FUNCTION_BLOCK MGZ_IMC (* Extracted Composite Function Block Type *)
  (* Standard: 61499-2 *)
  (* Version 10/20/2026, lizar *)
  PACKAGE Main;
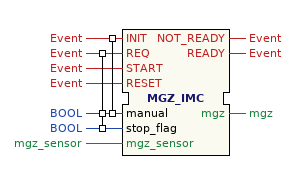
  EVENT_INPUT
    INIT WITH manual; (* Initialization Request *)
    REQ WITH manual, stop_flag; (* Normal Execution Request *)
    START;
    RESET;
  END_EVENT
  EVENT_OUTPUT
    NOT_READY;
    READY;
  END_EVENT
  VAR_INPUT
    manual : BOOL;
    stop_flag : BOOL;
  END_VAR
  SOCKETS
    mgz_sensor : mgz_sensor;
  END_SOCKETS
  PLUGS
    mgz : mgz;
  END_PLUGS
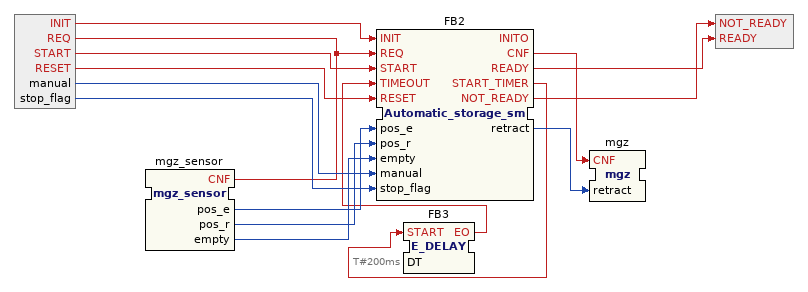
  FBS
    FB2 : Automatic_storage_sm;
    FB3 : E_DELAY(DT := T#200ms);
  END_FBS
  EVENT_CONNECTIONS
    FB2.START_TIMER TO FB3.START;
    FB3.EO TO FB2.TIMEOUT;
    INIT TO FB2.INIT;
    REQ TO FB2.REQ;
    START TO FB2.START;
    FB2.NOT_READY TO NOT_READY;
    FB2.READY TO READY;
    RESET TO FB2.RESET;
    FB2.CNF TO mgz.CNF;
    mgz_sensor.CNF TO FB2.REQ;
  END_CONNECTIONS
  DATA_CONNECTIONS
    manual TO FB2.manual;
    stop_flag TO FB2.stop_flag;
    FB2.retract TO mgz.retract;
    mgz_sensor.pos_e TO FB2.pos_e;
    mgz_sensor.pos_r TO FB2.pos_r;
    mgz_sensor.empty TO FB2.empty;
  END_CONNECTIONS
END_FUNCTION_BLOCK
